Fanuc KAREL source: kt00090.KL

-- PROVISIONAL review KL for V940-1; original PC SHA256 a83671e0cbe399e0cc62047c7a10c4224a22bcac312d8c066d9ed9cb463bd5e9
-- Incomplete behavior may be omitted. Consult companion uncertainty JSON. Do not deploy.
PROGRAM KT00090
%NOLOCKGROUP
VAR
  I2 : INTEGER
  OUT : REAL
-- UNRESOLVED_DECL H1 type=002017
BEGIN
  -- V9_ZERO_TABLE_METADATA_HINT layout=0001; no indexed target words; source/name/runtime held
  -- UNRESOLVED_PC offsets 5-19; opcodes 2E,22,9D,33,B4
  -- UNRESOLVED_PC offsets 24-35; opcodes 2E,23
  -- UNRESOLVED_PC offsets 40-63; opcodes 22,9D,33,B3,21,54,64,23
  -- UNRESOLVED_PC offsets 68-72; opcodes 7F
END KT00090
